(* IEC 61131-3 sources: rusty/compiler/plc_cfc/fixtures/blocks/valid/method_program, 1 file *)

(* ---- P.st ---- *)
PROGRAM P
VAR
    total : DINT;
END_VAR
METHOD bump : DINT
VAR_INPUT
    step : DINT;
END_VAR
    total := total + step;
    bump := total;
END_METHOD
END_PROGRAM
